// TIA Portal V21 export
TextList "TL_BalMode"  ListRange=Decimal
  TextListEntry   Text="0 lijevo/desno"
  TextListEntry   From=1, To=1, Text="1 + pramac/krma"
